// TIA Portal project "Camera" (V18)

(* hardware
DEVICE "S7-1200 station_1"  S7-1200 Station
   slot 0: "Rack_0"  S7-1200 Rack  Rack  V1.0
   slot 1: "PLC_1"  CPU 1215C DC/DC/DC  6ES7 215-1AG40-0XB0  V4.6
   slot 2: "SM 1278_1"  4SI IO link  6ES7 278-4BD32-0XB0  V2.1
   slot 3: "DI 2/DQ 2x24VDC_1"  DI2/DQ2 signal board  6ES7 223-0BD30-0XB0  V1.0
DEVICE "GSD device_1"  GSD.Device.PN
   slot 0: "Rack"  Rack  V1.0
   slot 0: "vos"  default module, no PDEV  VOSxxxx-F22x  V1.8
      slot 0: "default module, no PDEV"  default module, no PDEV
      slot 1: "input module 254 byte_1"  input module 254 byte
         slot 0: "input module 254 byte"  input module 254 byte
      slot 1: "Interface"  Interface
         slot 1: "Port 1"  Port 1
      slot 2: "output module 254 byte_1"  output module 254 byte
         slot 0: "output module 254 byte"  output module 254 byte
*)

// ===== PLC "PLC_1"  CPU 1215C DC/DC/DC =====

VAR_GLOBAL   // PLC tag table "Default tag table"
   "capteur 1" AT %I1.3 : Bool;
   "capteur 2" AT %I0.0 : Bool;
   "capteur 3" AT %I1.4 : Bool;
   "Km 1" AT %Q1.0 : Bool;
   "on" AT %I4.0 : Bool;
   "off" AT %I4.1 : Bool;
   "etape 0" AT %M1.0 : Bool;
   "etape 1" AT %M1.1 : Bool;
   "etape 2" AT %M1.2 : Bool;
   "etape 3" AT %M1.3 : Bool;
   "finT" AT %M1.4 : Bool;
   "Led" AT %Q0.0 : Bool;
END_VAR

// folder: System blocks/Program resources

DATA_BLOCK "IEC_Timer_0_DB"   // DB1
{ S7_Optimized_Access := 'TRUE' }
AUTHOR : Simatic
FAMILY : IEC
NAME : IEC_TMR
VERSION : 1.0
// stored: InstanceOfName IEC_TIMER
"IEC_TIMER"
BEGIN
END_DATA_BLOCK

// folder: (top level)

FUNCTION "sys" : Void   // FC1, LAD
{ S7_Optimized_Access := 'TRUE' }
VERSION : 0.1
BEGIN

REGION Network 2
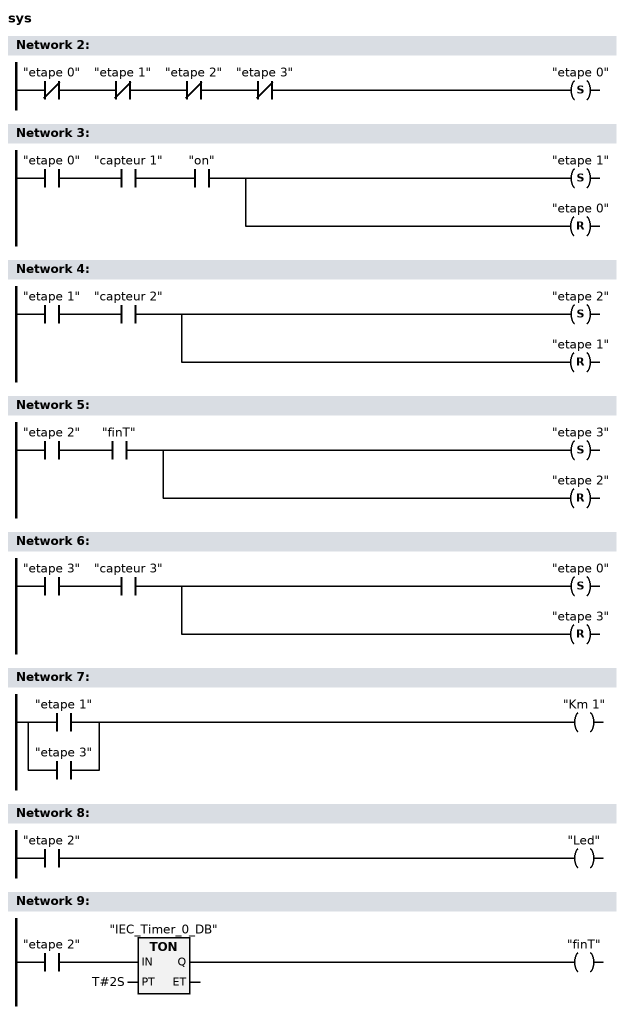
   RUNG wire#powerrail
      I_Contact( "etape 0" )
      I_Contact( "etape 1" )
      I_Contact( "etape 2" )
      I_Contact( "etape 3" )
      S_Coil( "etape 0" )
   END_RUNG
   // the same network as SCL:
   IF NOT "etape 0" AND NOT "etape 1" AND NOT "etape 2" AND NOT "etape 3" THEN "etape 0" := TRUE; END_IF;
END_REGION

REGION Network 3
   RUNG wire#powerrail
      Contact( "etape 0" )
      Contact( "capteur 1" )
      Contact( "on" )
      wire#w1
      S_Coil( "etape 1" )
   END_RUNG
   RUNG wire#w1
      R_Coil( "etape 0" )
   END_RUNG
   // the same network as SCL:
   IF "etape 0" AND "capteur 1" AND "on" THEN
       "etape 1" := TRUE;
       "etape 0" := FALSE;
   END_IF;
END_REGION

REGION Network 4
   RUNG wire#powerrail
      Contact( "etape 1" )
      Contact( "capteur 2" )
      wire#w1
      S_Coil( "etape 2" )
   END_RUNG
   RUNG wire#w1
      R_Coil( "etape 1" )
   END_RUNG
   // the same network as SCL:
   IF "etape 1" AND "capteur 2" THEN
       "etape 2" := TRUE;
       "etape 1" := FALSE;
   END_IF;
END_REGION

REGION Network 5
   RUNG wire#powerrail
      Contact( "etape 2" )
      Contact( "finT" )
      wire#w1
      S_Coil( "etape 3" )
   END_RUNG
   RUNG wire#w1
      R_Coil( "etape 2" )
   END_RUNG
   // the same network as SCL:
   IF "etape 2" AND "finT" THEN
       "etape 3" := TRUE;
       "etape 2" := FALSE;
   END_IF;
END_REGION

REGION Network 6
   RUNG wire#powerrail
      Contact( "etape 3" )
      Contact( "capteur 3" )
      wire#w1
      S_Coil( "etape 0" )
   END_RUNG
   RUNG wire#w1
      R_Coil( "etape 3" )
   END_RUNG
   // the same network as SCL:
   IF "etape 3" AND "capteur 3" THEN
       "etape 0" := TRUE;
       "etape 3" := FALSE;
   END_IF;
END_REGION

REGION Network 7
   RUNG wire#powerrail
      Contact( "etape 1" )
      wire#w1
      Coil( "Km 1" )
   END_RUNG
   RUNG wire#powerrail
      Contact( "etape 3" )
   END_RUNG wire#w1
   // the same network as SCL:
   "Km 1" := "etape 1" OR "etape 3";
END_REGION

REGION Network 8
   RUNG wire#powerrail
      Contact( "etape 2" )
      Coil( "Led" )
   END_RUNG
   // the same network as SCL:
   "Led" := "etape 2";
END_REGION

REGION Network 9
   "IEC_Timer_0_DB".TON(IN := "etape 2", PT := T#2S);
   "finT" := "IEC_Timer_0_DB".Q;
END_REGION
END_FUNCTION

FUNCTION "Led ctr" : Void   // FC2, LAD
{ S7_Optimized_Access := 'TRUE' }
VERSION : 0.1
BEGIN

REGION Network 1
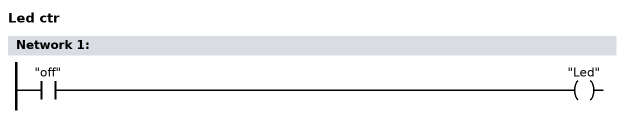
   RUNG wire#powerrail
      Contact( "off" )
      Coil( "Led" )
   END_RUNG
   // the same network as SCL:
   "Led" := "off";
END_REGION
END_FUNCTION

ORGANIZATION_BLOCK "Main"   // OB1, LAD, ProgramCycle
TITLE = "Main Program Sweep (Cycle)"
{ S7_Optimized_Access := 'TRUE' }
VERSION : 0.1
   VAR_INPUT
      Initial_Call : Bool;   // Initial call of this OB
      Remanence : Bool;   // =True, if remanent data are available
   END_VAR
BEGIN

REGION Network 1
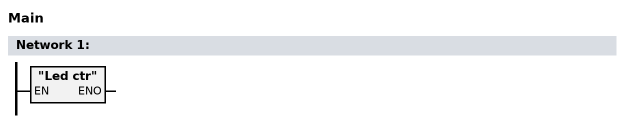
   RUNG wire#powerrail
      "Led ctr"()
   END_RUNG
   // the same network as SCL:
   "Led ctr"();
END_REGION
END_ORGANIZATION_BLOCK